TYPE E_LightAction :
(
    None,
    Toggle,
    TurnOn,
    TurnOff,
    SetBrightness
);
END_TYPE

(* stored: Version 1.1.0.1, ProductVersion 3.1.4026.20
   DUT E_LightAction: Id {D7C9A3E1-6F42-4A8D-9B31-2C5E7F901001} *)
